FUNCTION F_OpcUaCreatePaths (* Creates a browse name and a nodeId for OPC UA communication *)
  (* Standard: 61499-2; Description: Copyright (c) 2026 Monika Wenger This program and the accompanying materials are made available under the terms of the Eclipse Public License 2.0 which is available at https://www.eclipse.org/legal/epl-2.0/ SPDX-License-Identifier: EPL-2.0 *)
  (* Version 3.0, 2026-10-14, Monika Wenger *)
  PACKAGE eclipse4diac::opcua;
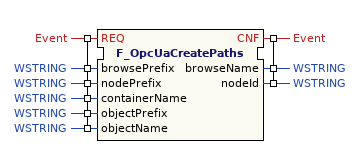
  EVENT_INPUT
    REQ WITH browsePrefix, nodePrefix, containerName, objectPrefix, objectName;
  END_EVENT
  EVENT_OUTPUT
    CNF WITH browseName, nodeId;
  END_EVENT
  VAR_INPUT
    browsePrefix : WSTRING;
    nodePrefix : WSTRING;
    containerName : WSTRING;
    objectPrefix : WSTRING;
    objectName : WSTRING;
  END_VAR
  VAR_OUTPUT
    browseName : WSTRING;
    nodeId : WSTRING;
  END_VAR
  BODY IN ST:
PACKAGE eclipse4diac::opcua;

(* Creates a browse name and a nodeId for OPC UA communication *)
FUNCTION F_OpcUaCreatePaths
VAR_INPUT
	browsePrefix : WSTRING;
	nodePrefix : WSTRING;
	containerName : WSTRING;
	objectPrefix : WSTRING;
	objectName : WSTRING;
END_VAR
VAR_OUTPUT
	browseName : WSTRING;
	nodeId : WSTRING;
END_VAR
VAR CONSTANT
	BROWSE_SEPARATOR : WSTRING := "/";
	NODE_SEPARATOR : WSTRING := ".";
END_VAR
IF EQ(objectPrefix, "") THEN
	browseName := CONCAT(browsePrefix, containerName, BROWSE_SEPARATOR, objectName);
	nodeId := CONCAT(nodePrefix, containerName, NODE_SEPARATOR, objectName);
ELSE
	browseName := CONCAT(browsePrefix, containerName, BROWSE_SEPARATOR, objectPrefix, BROWSE_SEPARATOR, objectName);
	nodeId := CONCAT(nodePrefix, containerName, NODE_SEPARATOR, objectPrefix, NODE_SEPARATOR, objectName);
END_IF;
END_FUNCTION
  END_BODY
END_FUNCTION
